(*
SPDX-FileCopyrightText: © 2026 Oleksandr Tiutyk <trofimich@gmail.com>
SPDX-License-Identifier: MIT
License: https://opensource.org/license/mit
*)

(*!
<summary>Selects the setup and outcome for a delayed timer observation.</summary>
*)

{attribute 'qualified_only'}
{attribute 'strict'}
TYPE DELAYED_TIMER_TEST_SCENARIO :
(
	//! <summary>Observe natural completion after delaying the first Execute.</summary>
	AFTER_START,
	//! <summary>Request cancellation after the preset but before any Execute.</summary>
	CANCEL_BEFORE_EXECUTE,
	//! <summary>Observe natural completion after restarting an active timer and delaying Execute.</summary>
	AFTER_ACTIVE_RESTART
);
END_TYPE

(* stored: Version 1.1.0.1
   DUT DELAYED_TIMER_TEST_SCENARIO: Id {f49a42df-8ee6-4ff9-a882-54c8b752cc82} *)
